ORGANIZATION_BLOCK "Cyclic 100mS"
TITLE = "Cyclic Interrupt"
VERSION : 0.1


VAR_TEMP
  OB35_EV_CLASS : BYTE ;	//Bits 0-3 = 1 (Coming event), Bits 4-7 = 1 (Event class 1)
  OB35_STRT_INF : BYTE ;	//16#36 (OB 35 has started)
  OB35_PRIORITY : BYTE ;	//Priority of OB Execution
  OB35_OB_NUMBR : BYTE ;	//35 (Organization block 35, OB35)
  OB35_RESERVED_1 : BYTE ;	//Reserved for system
  OB35_RESERVED_2 : BYTE ;	//Reserved for system
  OB35_PHASE_OFFSET : WORD ;	//Phase offset (msec)
  OB35_RESERVED_3 : INT ;	//Reserved for system
  OB35_EXC_FREQ : INT ;	//Frequency of execution (msec)
  OB35_DATE_TIME : DATE_AND_TIME ;	//Date and time OB35 started
END_VAR
BEGIN
NETWORK
TITLE =CYCLIC 100 mS

      CALL "GENERAL FAULTS" ;
      CALL "HMI CONTROL" ;
      CALL "HMI COMMS" ;
      CALL "LIGHT BAR" ;

//  CALL  "Sensor Check Calls"
NETWORK
TITLE =Lauer Comms

      CALL "LAUER CALL" ;

NETWORK
TITLE =Lauer Comms

      CALL "LAUER COMM FC" (
           UBDB                     := "DB LAUER",
           RXFA                     := 36,
           RXLE                     := 32,
           TXFA                     := 3,
           TXLE                     := 32,
           RSET                     := "M 210.1",
           TIMT                     := T    105,
           TIMZ                     := S5T#1S,
           COFF                     := "LAUER RESTART FC",
           INIT                     := "LAUER COMM ERR FC",
           RFLM                     := "M 210.0",
           EROR                     := "M 210.2");
END_ORGANIZATION_BLOCK
